FUNCTION_BLOCK EM_FbdCaller
VAR_INPUT
  ibInfeedClear : BOOL;
  ibSimulate    : BOOL;
END_VAR
VAR_OUTPUT
  obEmpty       : BOOL;
END_VAR
VAR
  fbLift        : CM_Lift;
END_VAR

// NETWORK 1

END_FUNCTION_BLOCK

(* stored: Version 1.1.0.1, ProductVersion 3.1.4024.12
   POU EM_FbdCaller: Id {0a1b2c3d-0000-4000-8000-000000000101}, SpecialFunc None *)
